Staubli VAL3: utText.dtx

public string sFontFamily
public string sFontStyle
public string sFontWeight
public string sTextAlignment
public num nFontSize
